(* IEC 61131-3 sources: plc-st-coding-agent/progress/evidence/v13_rescore_20261108/candidates/codex_minimax-m27, 19 files *)

(* ---- public-easy-01.st ---- *)
FUNCTION_BLOCK FB
VAR_INPUT
    bottleSensor           : BOOL;
    cleaningConfirmButton  : BOOL;
    fillingConfirmButton   : BOOL;
    cappingConfirmButton   : BOOL;
    packingConfirmButton   : BOOL;
    finishedButton         : BOOL;
END_VAR

VAR_OUTPUT
    Pump_Motor        : BOOL;
    Filling_Valve     : BOOL;
    Capping_Machine   : BOOL;
    Packing_Machine   : BOOL;
    Completion_Light  : BOOL;
END_VAR

VAR
    step                  : INT := 0;
    prevBottleSensor      : BOOL := FALSE;
    prevCleaningConfirm   : BOOL := FALSE;
    prevFillingConfirm    : BOOL := FALSE;
    prevCappingConfirm    : BOOL := FALSE;
    prevPackingConfirm    : BOOL := FALSE;
    prevFinishedButton    : BOOL := FALSE;
END_VAR

// Rising edge detection
VAR
    bottleRising         : BOOL;
    cleaningRising       : BOOL;
    fillingRising        : BOOL;
    cappingRising        : BOOL;
    packingRising        : BOOL;
    finishedRising       : BOOL;
END_VAR

bottleRising       := bottleSensor        AND NOT prevBottleSensor;
cleaningRising     := cleaningConfirmButton  AND NOT prevCleaningConfirm;
fillingRising      := fillingConfirmButton   AND NOT prevFillingConfirm;
cappingRising      := cappingConfirmButton   AND NOT prevCappingConfirm;
packingRising      := packingConfirmButton   AND NOT prevPackingConfirm;
finishedRising     := finishedButton      AND NOT prevFinishedButton;

// State machine transitions
IF step = 0 THEN
    IF bottleRising THEN
        step := 1;
    END_IF
ELSIF step = 1 THEN
    IF cleaningRising THEN
        step := 2;
    END_IF
ELSIF step = 2 THEN
    IF fillingRising THEN
        step := 3;
    END_IF
ELSIF step = 3 THEN
    IF cappingRising THEN
        step := 4;
    END_IF
ELSIF step = 4 THEN
    IF packingRising THEN
        step := 5;
    END_IF
END_IF

// Output logic based on step
Pump_Motor       := (step >= 1);
Filling_Valve    := (step >= 2);
Capping_Machine  := (step >= 3);
Packing_Machine  := (step >= 4);
Completion_Light := (step >= 5);

// Reset on finishedButton rising only when in COMPLETE state
IF finishedRising AND (step = 5) THEN
    step := 0;
END_IF

// Update previous states
prevBottleSensor    := bottleSensor;
prevCleaningConfirm := cleaningConfirmButton;
prevFillingConfirm  := fillingConfirmButton;
prevCappingConfirm  := cappingConfirmButton;
prevPackingConfirm  := packingConfirmButton;
prevFinishedButton  := finishedButton;
END_FUNCTION_BLOCK

(* ---- public-easy-02.st ---- *)
FUNCTION_BLOCK FB
VAR_INPUT
END_VAR
VAR_OUTPUT
    hasChanged      : BOOL;
    hasRisingEdges  : BOOL;
    risingBits      : DWORD;
    noOfRisingBits  : USINT;
    hasFallingEdges : BOOL;
    fallingBits     : DWORD;
    noOfFallingBits : USINT;
END_VAR
VAR
    prevValue : DWORD := 0;
    bitCheck  : DWORD;
    i         : USINT;
END_VAR

// Calculate rising edges: current=1 AND previous=0
risingBits := value AND NOT prevValue;

// Calculate falling edges: current=0 AND previous=1
fallingBits := NOT value AND prevValue;

// Detect if value has changed
hasChanged := (value <> prevValue);

// Set edge flags based on bit streams
hasRisingEdges := (risingBits <> 0);
hasFallingEdges := (fallingBits <> 0);

// Count rising bits
noOfRisingBits := 0;
bitCheck := risingBits;
FOR i := 0 TO 31 DO
    IF (bitCheck AND 1) = 1 THEN
        noOfRisingBits := noOfRisingBits + 1;
    END_IF;
    bitCheck := SHR(bitCheck, 1);
END_FOR;

// Count falling bits
noOfFallingBits := 0;
bitCheck := fallingBits;
FOR i := 0 TO 31 DO
    IF (bitCheck AND 1) = 1 THEN
        noOfFallingBits := noOfFallingBits + 1;
    END_IF;
    bitCheck := SHR(bitCheck, 1);
END_FOR;

// Update history for next cycle
prevValue := value;
END_FUNCTION_BLOCK

(* ---- public-easy-03.st ---- *)
FUNCTION_BLOCK FB
VAR_INPUT
    Value       : REAL;
    hiLevel     : REAL;
    loLevel     : REAL;
    hystWindow  : REAL;
END_VAR
VAR_OUTPUT
    hiAlarm     : BOOL;
    loAlarm     : BOOL;
    error       : BOOL;
    status      : WORD;
END_VAR

    // Parameter validation errors take priority
    IF loLevel >= hiLevel THEN
        error   := TRUE;
        status  := 16#8001;
        RETURN;
    END_IF

    IF hystWindow >= (hiLevel - loLevel) THEN
        error   := TRUE;
        status  := 16#8002;
        RETURN;
    END_IF

    // No error
    error  := FALSE;
    status := 16#0000;

    // High alarm with hysteresis
    // Trigger: Value > hiLevel
    // Reset:   Value < hiLevel - hystWindow
    IF Value > hiLevel THEN
        hiAlarm := TRUE;
    ELSIF Value < (hiLevel - hystWindow) THEN
        hiAlarm := FALSE;
    END_IF

    // Low alarm with hysteresis
    // Trigger: Value < loLevel
    // Reset:   Value > loLevel + hystWindow
    IF Value < loLevel THEN
        loAlarm := TRUE;
    ELSIF Value > (loLevel + hystWindow) THEN
        loAlarm := FALSE;
    END_IF

END_FUNCTION_BLOCK

(* ---- public-easy-04.st ---- *)
FUNCTION_BLOCK FB
VAR_INPUT
    VISCOSITY_OK     : BOOL;
    PASTE_E_STOP_NC  : BOOL;
    DebounceTime     : TIME;
    CycleTime        : TIME;
END_VAR
VAR_OUTPUT
    VFD_RUN          : BOOL;
    PUMP_MAINT_DUE   : BOOL;
    PUMP_RUNTIME_ACC : LINT;
END_VAR
VAR
    visc_debounce_acc : TIME := T#0s;
    visc_valid        : BOOL := FALSE;
END_VAR

// Debounce logic for viscosity condition
IF NOT VISCOSITY_OK THEN
    visc_debounce_acc := T#0s;
    visc_valid        := FALSE;
ELSIF visc_debounce_acc < DebounceTime THEN
    visc_debounce_acc := visc_debounce_acc + CycleTime;
    IF visc_debounce_acc >= DebounceTime THEN
        visc_debounce_acc := DebounceTime;
        visc_valid        := TRUE;
    END_IF
END_IF;

// VFD run permissive: E-STOP must be closed AND viscosity debounced valid
VFD_RUN := PASTE_E_STOP_NC AND visc_valid;

// Accumulate runtime (in hours) only while pump is running
IF VFD_RUN THEN
    PUMP_RUNTIME_ACC := PUMP_RUNTIME_ACC + TO_LINT(TIME_TO_INT(CycleTime) / 3600000);
END_IF;

// Maintenance due indication at 500 hours
PUMP_MAINT_DUE := (PUMP_RUNTIME_ACC >= 500);
END_FUNCTION_BLOCK

(* ---- public-easy-05.st ---- *)
FUNCTION_BLOCK FB
VAR_INPUT
    Gap_Exceeded : BOOL;
    Weld_E_Stop_NC : BOOL;
    DebounceTime : TIME;
END_VAR
VAR_OUTPUT
    Operator_Alert : BOOL;
    Weld_Soft_Start_Active : BOOL;
END_VAR
VAR
    init_cycle_count : INT := 5;
    gap_exceeded_prev : BOOL := FALSE;
    debounce_counter : INT := 0;
    debounce_required : INT := 50;
END_VAR

// Emergency stop priority - immediate reset regardless of state
IF NOT Weld_E_Stop_NC THEN
    Operator_Alert := FALSE;
    debounce_counter := 0;
    Weld_Soft_Start_Active := FALSE;
    gap_exceeded_prev := Gap_Exceeded;
    RETURN;
END_IF;

// Power-up initialization inhibition (5 scan cycles)
IF init_cycle_count > 0 THEN
    init_cycle_count := init_cycle_count - 1;
    Weld_Soft_Start_Active := TRUE;
    Operator_Alert := FALSE;
    debounce_counter := 0;
    gap_exceeded_prev := Gap_Exceeded;
    RETURN;
END_IF;

Weld_Soft_Start_Active := FALSE;
gap_exceeded_prev := Gap_Exceeded;

// Gap monitoring with debounce
IF Gap_Exceeded THEN
    debounce_counter := debounce_counter + 1;
    IF debounce_counter >= debounce_required THEN
        Operator_Alert := TRUE;
    ELSE
        Operator_Alert := FALSE;
    END_IF;
ELSE
    debounce_counter := 0;
    Operator_Alert := FALSE;
END_IF;
END_FUNCTION_BLOCK

(* ---- public-easy-06.st ---- *)
FUNCTION_BLOCK FB
VAR_INPUT
    DO_LOW : BOOL;
    AERATION_E_STOP_NC : BOOL;
END_VAR
VAR_OUTPUT
    BLOWER_RUN : BOOL;
    AERATION_BLOWER_CYCLE_COUNT : UINT;
END_VAR
VAR
    prev_blower_run : BOOL := FALSE;
    delay_counter : UINT := 0;
END_VAR

IF DO_LOW AND AERATION_E_STOP_NC THEN
    IF delay_counter < 5 THEN
        delay_counter := delay_counter + 1;
    END_IF
    IF delay_counter >= 5 THEN
        BLOWER_RUN := TRUE;
    ELSE
        BLOWER_RUN := FALSE;
    END_IF
ELSE
    BLOWER_RUN := FALSE;
    delay_counter := 0;
END_IF

IF BLOWER_RUN AND NOT prev_blower_run THEN
    AERATION_BLOWER_CYCLE_COUNT := AERATION_BLOWER_CYCLE_COUNT + 1;
END_IF

prev_blower_run := BLOWER_RUN;
END_FUNCTION_BLOCK

(* ---- public-hard-01.st ---- *)
FUNCTION_BLOCK FB
VAR_INPUT
    estop            : BOOL;
    opeMode          : BOOL;
    valveAStart      : BOOL;
    valveBStart      : BOOL;
    valveCStart      : BOOL;
    valveDStart      : BOOL;
    mixMotorStart    : BOOL;
    autoStart        : BOOL;
    processMode      : BOOL;
    levelSensor      : INT;
    mixMotorComplete : BOOL;
END_VAR
VAR_OUTPUT
    valveARun    : BOOL;
    valveBRun    : BOOL;
    valveCRun    : BOOL;
    valveDRun    : BOOL;
    mixMotorRun  : BOOL;
END_VAR
VAR
    // Auto mode state machine
    autoState : INT;
    // Rising edge detection history
    prevValveAStart    : BOOL;
    prevValveBStart    : BOOL;
    prevValveCStart    : BOOL;
    prevValveDStart    : BOOL;
    prevMixMotorStart  : BOOL;
    prevAutoStart      : BOOL;
    // Rising edge results
    valveAStartEdge    : BOOL;
    valveBStartEdge    : BOOL;
    valveCStartEdge    : BOOL;
    valveDStartEdge    : BOOL;
    mixMotorStartEdge  : BOOL;
    autoStartEdge      : BOOL;
END_VAR

    // Auto state constants
    // 0=IDLE, 1=VALVE_A, 2=VALVE_B, 3=VALVE_C, 4=MIXING, 5=DISCHARGE

    // Rising edge detection
    valveAStartEdge   := valveAStart AND NOT prevValveAStart;
    valveBStartEdge   := valveBStart AND NOT prevValveBStart;
    valveCStartEdge   := valveCStart AND NOT prevValveCStart;
    valveDStartEdge   := valveDStart AND NOT prevValveDStart;
    mixMotorStartEdge := mixMotorStart AND NOT prevMixMotorStart;
    autoStartEdge     := autoStart AND NOT prevAutoStart;

    // Update edge detection history
    prevValveAStart   := valveAStart;
    prevValveBStart   := valveBStart;
    prevValveCStart   := valveCStart;
    prevValveDStart   := valveDStart;
    prevMixMotorStart := mixMotorStart;
    prevAutoStart     := autoStart;

    // Default outputs off (safety)
    valveARun   := FALSE;
    valveBRun   := FALSE;
    valveCRun   := FALSE;
    valveDRun   := FALSE;
    mixMotorRun := FALSE;

    // Emergency stop - all equipment stops immediately
    IF NOT estop THEN
        autoState := 0;
        RETURN;
    END_IF

    // Manual mode
    IF NOT opeMode THEN
        // Rising edge toggles for each device
        IF valveAStartEdge THEN
            valveARun := NOT valveARun;
        END_IF
        IF valveBStartEdge THEN
            valveBRun := NOT valveBRun;
        END_IF
        IF valveCStartEdge THEN
            valveCRun := NOT valveCRun;
        END_IF
        IF valveDStartEdge THEN
            valveDRun := NOT valveDRun;
        END_IF
        IF mixMotorStartEdge THEN
            mixMotorRun := NOT mixMotorRun;
        END_IF
    // Automatic mode
    ELSIF opeMode THEN
        CASE autoState OF
            0: // IDLE
                IF autoStartEdge THEN
                    autoState := 1;
                END_IF

            1: // Open Valve A
                valveARun := TRUE;
                IF levelSensor >= 50 THEN
                    valveARun := FALSE;
                    autoState := 2;
                END_IF

            2: // Open Valve B
                valveBRun := TRUE;
                IF levelSensor >= 80 THEN
                    valveBRun := FALSE;
                    IF processMode THEN
                        autoState := 3;
                    ELSE
                        autoState := 4;
                    END_IF;
                END_IF

            3: // Open Valve C (processMode=true)
                valveCRun := TRUE;
                IF levelSensor >= 100 THEN
                    valveCRun := FALSE;
                    autoState := 4;
                END_IF

            4: // Mixing
                mixMotorRun := TRUE;
                IF mixMotorComplete THEN
                    mixMotorRun := FALSE;
                    autoState := 5;
                END_IF

            5: // Discharge through Valve D
                valveDRun := TRUE;
                IF levelSensor <= 0 THEN
                    valveDRun := FALSE;
                    autoState := 0;
                END_IF
        END_CASE
    END_IF

END_FUNCTION_BLOCK

(* ---- public-hard-02.st ---- *)
FUNCTION_BLOCK FB
VAR_INPUT
    processLength : USINT;
    sensor1 : BOOL;
    sensor2 : BOOL;
    sensor3 : BOOL;
    sensor4 : BOOL;
    sensor5 : BOOL;
    station1Start : BOOL;
    station2Complete : BOOL;
    station3Complete : BOOL;
    station4Complete : BOOL;
    processSequence : ARRAY[1..8] OF USINT;
END_VAR

VAR_OUTPUT
    conveyorLeft : BOOL;
    conveyorRight : BOOL;
END_VAR

VAR
    phase : USINT := 0;
    curStation : USINT := 0;
    dstStation : USINT := 0;
    idx : USINT := 1;
    prevStart : BOOL := FALSE;
    prevComp2 : BOOL := FALSE;
    prevComp3 : BOOL := FALSE;
    prevComp4 : BOOL := FALSE;
END_VAR

VAR
    startEdge : BOOL;
    compEdge : BOOL;
END_VAR

startEdge := station1Start AND NOT prevStart;
compEdge := (station2Complete AND NOT prevComp2) OR
            (station3Complete AND NOT prevComp3) OR
            (station4Complete AND NOT prevComp4);

prevStart := station1Start;
prevComp2 := station2Complete;
prevComp3 := station3Complete;
prevComp4 := station4Complete;

IF sensor1 AND startEdge THEN
    phase := 0;
    idx := 1;
    curStation := 1;
END_IF

CASE phase OF
    0:
        conveyorLeft := FALSE;
        conveyorRight := FALSE;
        IF sensor1 AND startEdge THEN
            curStation := 1;
            idx := 1;
            dstStation := processSequence[idx];
            phase := 1;
        END_IF

    1:
        IF dstStation > curStation THEN
            conveyorRight := TRUE;
            conveyorLeft := FALSE;
        ELSIF dstStation < curStation THEN
            conveyorLeft := TRUE;
            conveyorRight := FALSE;
        END_IF

        IF (dstStation = 2 AND sensor2) OR
           (dstStation = 3 AND sensor3) OR
           (dstStation = 4 AND sensor4) OR
           (dstStation = 5 AND sensor5) THEN
            curStation := dstStation;
            conveyorLeft := FALSE;
            conveyorRight := FALSE;
            phase := 2;
        END_IF

    2:
        conveyorLeft := FALSE;
        conveyorRight := FALSE;

        IF compEdge THEN
            IF curStation = 2 THEN
                idx := idx + 1;
                IF idx <= processLength THEN
                    dstStation := processSequence[idx];
                    phase := 1;
                END_IF
            ELSIF curStation = 3 THEN
                idx := idx + 1;
                IF idx <= processLength THEN
                    dstStation := processSequence[idx];
                    phase := 1;
                END_IF
            ELSIF curStation = 4 THEN
                idx := idx + 1;
                IF idx <= processLength THEN
                    dstStation := processSequence[idx];
                    phase := 1;
                END_IF
            END_IF
        END_IF

        IF curStation = 5 THEN
            phase := 0;
        END_IF
END_CASE
END_FUNCTION_BLOCK

(* ---- public-hard-03.st ---- *)
TYPE ST_Recipe :
STRUCT
    recipeID : INT;
    ingredientType : INT;
    ingredientRatio : REAL;
    productionTemperature : REAL;
END_STRUCT
END_TYPE

FUNCTION_BLOCK FB
VAR_INPUT
    addRecipe : BOOL;
    deleteRecipe : BOOL;
    modifyRecipe : BOOL;
    queryRecipe : BOOL;
    recipeIn : ST_Recipe;
END_VAR

VAR_OUTPUT
    recipeAdded : BOOL := FALSE;
    recipeDeleted : BOOL := FALSE;
    recipeModified : BOOL := FALSE;
    recipeQueryResult : ST_Recipe;
    error : BOOL := FALSE;
    status : WORD := 16#0000;
END_VAR

VAR_IN_OUT
    recipe : ARRAY[1..10] OF ST_Recipe;
END_VAR

VAR
    addRecipePrev : BOOL := FALSE;
    deleteRecipePrev : BOOL := FALSE;
    modifyRecipePrev : BOOL := FALSE;
    queryRecipePrev : BOOL := FALSE;
    foundIndex : INT;
    i : INT;
    isDuplicate : BOOL;
    isFound : BOOL;
END_VAR

    error := FALSE;
    status := 16#0000;
    recipeAdded := FALSE;
    recipeDeleted := FALSE;
    recipeModified := FALSE;

    IF addRecipe AND NOT addRecipePrev THEN
        isDuplicate := FALSE;
        isFound := FALSE;
        foundIndex := 0;

        FOR i := 1 TO 10 DO
            IF recipe[i].recipeID = recipeIn.recipeID AND recipeIn.recipeID <> 0 THEN
                isDuplicate := TRUE;
                EXIT;
            END_IF
        END_FOR

        IF isDuplicate THEN
            error := TRUE;
            status := 16#8002;
        ELSE
            foundIndex := 0;
            FOR i := 1 TO 10 DO
                IF recipe[i].recipeID = 0 THEN
                    foundIndex := i;
                    EXIT;
                END_IF
            END_FOR

            IF foundIndex = 0 THEN
                error := TRUE;
                status := 16#8003;
            ELSE
                recipe[foundIndex] := recipeIn;
                recipeAdded := TRUE;
            END_IF
        END_IF
    END_IF

    IF deleteRecipe AND NOT deleteRecipePrev THEN
        isFound := FALSE;
        foundIndex := 0;

        FOR i := 1 TO 10 DO
            IF recipe[i].recipeID = recipeIn.recipeID AND recipeIn.recipeID <> 0 THEN
                isFound := TRUE;
                foundIndex := i;
                EXIT;
            END_IF
        END_FOR

        IF NOT isFound THEN
            error := TRUE;
            status := 16#8004;
        ELSE
            recipe[foundIndex].recipeID := 0;
            recipeDeleted := TRUE;
        END_IF
    END_IF

    IF modifyRecipe AND NOT modifyRecipePrev THEN
        isFound := FALSE;
        foundIndex := 0;

        FOR i := 1 TO 10 DO
            IF recipe[i].recipeID = recipeIn.recipeID AND recipeIn.recipeID <> 0 THEN
                isFound := TRUE;
                foundIndex := i;
                EXIT;
            END_IF
        END_FOR

        IF NOT isFound THEN
            error := TRUE;
            status := 16#8005;
        ELSE
            recipe[foundIndex] := recipeIn;
            recipeModified := TRUE;
        END_IF
    END_IF

    IF queryRecipe AND NOT queryRecipePrev THEN
        isFound := FALSE;
        foundIndex := 0;

        FOR i := 1 TO 10 DO
            IF recipe[i].recipeID = recipeIn.recipeID AND recipeIn.recipeID <> 0 THEN
                isFound := TRUE;
                foundIndex := i;
                EXIT;
            END_IF
        END_FOR

        IF NOT isFound THEN
            error := TRUE;
            status := 16#8001;
        ELSE
            recipeQueryResult := recipe[foundIndex];
        END_IF
    END_IF

    addRecipePrev := addRecipe;
    deleteRecipePrev := deleteRecipe;
    modifyRecipePrev := modifyRecipe;
    queryRecipePrev := queryRecipe;

END_FUNCTION_BLOCK

(* ---- public-hard-04.st ---- *)
FUNCTION_BLOCK FB
VAR_INPUT
    enqueue  : BOOL;
    dequeue  : BOOL;
    reset    : BOOL;
    capacity : DINT;
END_VAR
VAR_OUTPUT
    elementCount : DINT := 0;
    status       : WORD := 16#0000;
END_VAR
VAR_IN_OUT
    item   : DINT;
    buffer : ARRAY[1..4] OF DINT;
END_VAR
VAR
    head        : DINT := 1;
    tail        : DINT := 1;
    lastEnqueue : BOOL := FALSE;
    lastDequeue : BOOL := FALSE;
    lastReset   : BOOL := FALSE;
END_VAR

status := 16#0000;

IF reset THEN
    elementCount := 0;
    head := 1;
    tail := 1;
ELSIF NOT lastReset THEN
    IF enqueue AND NOT lastEnqueue THEN
        IF elementCount < capacity THEN
            buffer[tail] := item;
            elementCount := elementCount + 1;
            tail := (tail MOD capacity) + 1;
        ELSE
            status := 16#8002;
        END_IF
    ELSIF dequeue AND NOT lastDequeue THEN
        IF elementCount > 0 THEN
            item := buffer[head];
            elementCount := elementCount - 1;
            head := (head MOD capacity) + 1;
        ELSE
            status := 16#8001;
        END_IF
    END_IF
END_IF

lastEnqueue := enqueue;
lastDequeue := dequeue;
lastReset   := reset;
END_FUNCTION_BLOCK

(* ---- public-hard-05.st ---- *)
FUNCTION_BLOCK FB
VAR_INPUT
    ManualMode : BOOL;
    SingleStepMode : BOOL;
    SingleCycleMode : BOOL;
    ContinuousMode : BOOL;
    EmergencyStop : BOOL;
    Start : BOOL;
    DownButton : BOOL;
    UpButton : BOOL;
    LeftButton : BOOL;
    RightButton : BOOL;
    GripButton : BOOL;
    ReleaseButton : BOOL;
    DownLimitSwitch : BOOL;
    UpLimitSwitch : BOOL;
    LeftLimitSwitch : BOOL;
    RightLimitSwitch : BOOL;
    GripLimitSwitch : BOOL;
    ReleaseLimitSwitch : BOOL;
END_VAR

VAR_OUTPUT
    MoveDown : BOOL := FALSE;
    MoveUp : BOOL := FALSE;
    MoveLeft : BOOL := FALSE;
    MoveRight : BOOL := FALSE;
    ActivateGrip : BOOL := FALSE;
    ActivateRelease : BOOL := FALSE;
END_VAR

VAR
    Step : INT := 1;
    StartPrev : BOOL := FALSE;
    IsRunning : BOOL := FALSE;
END_VAR

    // Edge detection for Start button
    VAR
        StartRisingEdge : BOOL;
    END_VAR
    StartRisingEdge := Start AND NOT StartPrev;
    StartPrev := Start;

    // Emergency stop - highest priority
    IF NOT EmergencyStop THEN
        MoveDown := FALSE;
        MoveUp := FALSE;
        MoveLeft := FALSE;
        MoveRight := FALSE;
        ActivateGrip := FALSE;
        ActivateRelease := FALSE;
        RETURN;
    END_IF

    // Mode initialization
    IF SingleStepMode THEN
        IF NOT IsRunning THEN
            IF StartRisingEdge THEN
                Step := 1;
                IsRunning := TRUE;
            END_IF;
        END_IF;
    ELSIF SingleCycleMode THEN
        IF NOT IsRunning THEN
            IF StartRisingEdge THEN
                Step := 1;
                IsRunning := TRUE;
            END_IF;
        END_IF;
    ELSIF ContinuousMode THEN
        IF NOT IsRunning THEN
            IF StartRisingEdge THEN
                Step := 1;
                IsRunning := TRUE;
            END_IF;
        END_IF;
    ELSE
        IsRunning := FALSE;
    END_IF;

    // Execute current step in automatic modes
    IF IsRunning THEN
        CASE Step OF
            1: // MoveDown
                MoveDown := TRUE;
                IF DownLimitSwitch THEN
                    MoveDown := FALSE;
                    IF Step < 8 THEN
                        Step := Step + 1;
                    ELSE
                        Step := 1;
                    END_IF;
                    IF SingleStepMode THEN
                        IsRunning := FALSE;
                    END_IF;
                END_IF;

            2: // ActivateGrip
                ActivateGrip := TRUE;
                IF GripLimitSwitch THEN
                    ActivateGrip := FALSE;
                    IF Step < 8 THEN
                        Step := Step + 1;
                    ELSE
                        Step := 1;
                    END_IF;
                    IF SingleStepMode THEN
                        IsRunning := FALSE;
                    END_IF;
                END_IF;

            3: // MoveUp
                MoveUp := TRUE;
                IF UpLimitSwitch THEN
                    MoveUp := FALSE;
                    IF Step < 8 THEN
                        Step := Step + 1;
                    ELSE
                        Step := 1;
                    END_IF;
                    IF SingleStepMode THEN
                        IsRunning := FALSE;
                    END_IF;
                END_IF;

            4: // MoveRight
                MoveRight := TRUE;
                IF RightLimitSwitch THEN
                    MoveRight := FALSE;
                    IF Step < 8 THEN
                        Step := Step + 1;
                    ELSE
                        Step := 1;
                    END_IF;
                    IF SingleStepMode THEN
                        IsRunning := FALSE;
                    END_IF;
                END_IF;

            5: // MoveDown
                MoveDown := TRUE;
                IF DownLimitSwitch THEN
                    MoveDown := FALSE;
                    IF Step < 8 THEN
                        Step := Step + 1;
                    ELSE
                        Step := 1;
                    END_IF;
                    IF SingleStepMode THEN
                        IsRunning := FALSE;
                    END_IF;
                END_IF;

            6: // ActivateRelease
                ActivateRelease := TRUE;
                IF ReleaseLimitSwitch THEN
                    ActivateRelease := FALSE;
                    IF Step < 8 THEN
                        Step := Step + 1;
                    ELSE
                        Step := 1;
                    END_IF;
                    IF SingleStepMode THEN
                        IsRunning := FALSE;
                    END_IF;
                END_IF;

            7: // MoveUp
                MoveUp := TRUE;
                IF UpLimitSwitch THEN
                    MoveUp := FALSE;
                    IF Step < 8 THEN
                        Step := Step + 1;
                    ELSE
                        Step := 1;
                    END_IF;
                    IF SingleStepMode THEN
                        IsRunning := FALSE;
                    END_IF;
                END_IF;

            8: // MoveLeft
                MoveLeft := TRUE;
                IF LeftLimitSwitch THEN
                    MoveLeft := FALSE;
                    Step := 1;
                    IF SingleStepMode THEN
                        IsRunning := FALSE;
                    END_IF;
                END_IF;
        END_CASE;

    // Manual mode
    ELSIF ManualMode THEN
        // Down
        MoveDown := DownButton AND NOT DownLimitSwitch;
        // Up
        MoveUp := UpButton AND NOT UpLimitSwitch;
        // Left
        MoveLeft := LeftButton AND NOT LeftLimitSwitch;
        // Right
        MoveRight := RightButton AND NOT RightLimitSwitch;
        // Grip
        ActivateGrip := GripButton AND NOT GripLimitSwitch;
        // Release
        ActivateRelease := ReleaseButton AND NOT ReleaseLimitSwitch;
    END_IF;

END_FUNCTION_BLOCK

(* ---- public-hard-06.st ---- *)
FUNCTION_BLOCK FB
VAR_INPUT
    Mode            : BOOL;
    ForwardButton   : BOOL;
    ReverseButton   : BOOL;
    SensorFeed      : BOOL;
    SensorWash      : BOOL;
    SensorWeight    : BOOL;
    SensorFiring    : BOOL;
    SensorOutput    : BOOL;
    washComplete    : BOOL;
    weightComplete  : BOOL;
    weight          : REAL;
    firingComplete  : BOOL;
END_VAR
VAR_OUTPUT
    MotorForward    : BOOL;
    MotorReverse    : BOOL;
    kick            : BOOL;
    CompletionLight : BOOL;
    firingTemp      : REAL;
END_VAR
VAR
    eState              : INT;
    prevForwardButton   : BOOL;
    prevReverseButton   : BOOL;
    prevwashComplete    : BOOL;
    prevweightComplete  : BOOL;
    prevfiringComplete  : BOOL;
    bKickDone           : BOOL;
END_VAR

    // Edge detection: rising edge flags
    VAR
        bFwdRising   : BOOL;
        bRevRising   : BOOL;
        bWashRising  : BOOL;
        bWeightRising: BOOL;
        bFiringRising: BOOL;
    END_VAR

    bFwdRising   := (NOT prevForwardButton)  AND ForwardButton;
    bRevRising   := (NOT prevReverseButton)  AND ReverseButton;
    bWashRising  := (NOT prevwashComplete)   AND washComplete;
    bWeightRising:= (NOT prevweightComplete) AND weightComplete;
    bFiringRising:= (NOT prevfiringComplete) AND firingComplete;

    // Reset kick flag on new cycle start (ForwardButton rising edge in any mode)
    IF bFwdRising THEN
        bKickDone := FALSE;
    END_IF

    IF Mode = FALSE THEN
        // Manual mode
        eState := 0;
        MotorForward := ForwardButton;
        MotorReverse := ReverseButton;
        kick := FALSE;
        CompletionLight := FALSE;
        firingTemp := 0.0;
    ELSE
        // Automatic mode
        CASE eState OF
            0:  // IDLE
                MotorForward := FALSE;
                MotorReverse := FALSE;
                kick := FALSE;
                CompletionLight := FALSE;
                firingTemp := 0.0;
                bKickDone := FALSE;
                IF SensorFeed THEN
                    eState := 1;
                END_IF

            1:  // MOVING_TO_WASH
                MotorForward := TRUE;
                MotorReverse := FALSE;
                kick := FALSE;
                IF SensorWash THEN
                    eState := 2;
                END_IF

            2:  // AT_WASH
                MotorForward := FALSE;
                MotorReverse := FALSE;
                kick := FALSE;
                IF bWashRising THEN
                    eState := 3;
                END_IF

            3:  // MOVING_TO_WEIGH
                MotorForward := TRUE;
                MotorReverse := FALSE;
                kick := FALSE;
                IF SensorWeight THEN
                    eState := 4;
                END_IF

            4:  // AT_WEIGH
                MotorForward := FALSE;
                MotorReverse := FALSE;
                kick := FALSE;
                IF bWeightRising THEN
                    IF weight >= 100.0 AND weight <= 200.0 THEN
                        firingTemp := 500.0 + (weight - 100.0) * 0.5;
                        eState := 6;
                    ELSE
                        eState := 5;
                    END_IF;
                END_IF

            5:  // KICKING
                MotorForward := FALSE;
                MotorReverse := FALSE;
                kick := TRUE;
                IF NOT bKickDone THEN
                    bKickDone := TRUE;
                    eState := 0;
                END_IF

            6:  // MOVING_TO_FIRING
                MotorForward := TRUE;
                MotorReverse := FALSE;
                kick := FALSE;
                IF SensorFiring THEN
                    eState := 7;
                END_IF

            7:  // AT_FIRING
                MotorForward := FALSE;
                MotorReverse := FALSE;
                kick := FALSE;
                IF bFiringRising THEN
                    eState := 8;
                END_IF

            8:  // MOVING_TO_OUTPUT
                MotorForward := TRUE;
                MotorReverse := FALSE;
                kick := FALSE;
                IF SensorOutput THEN
                    eState := 9;
                END_IF

            9:  // AT_OUTPUT
                MotorForward := FALSE;
                MotorReverse := FALSE;
                kick := FALSE;
                CompletionLight := SensorOutput;
                IF NOT SensorOutput THEN
                    eState := 0;
                END_IF

        END_CASE
    END_IF

    prevForwardButton  := ForwardButton;
    prevReverseButton  := ReverseButton;
    prevwashComplete   := washComplete;
    prevweightComplete := weightComplete;
    prevfiringComplete := firingComplete;

END_FUNCTION_BLOCK

(* ---- public-medium-01.st ---- *)
TYPE ST_Pump
    STRUCT
        priority   : INT;
        selection  : BOOL;
        RunComd    : BOOL;
    END_STRUCT
END_TYPE

FUNCTION_BLOCK FB
VAR_INPUT
    mode  : BOOL;
    start : BOOL;
    stop  : BOOL;
END_VAR
VAR_IN_OUT
    pumpGroup : ARRAY[1..5] OF ST_Pump;
END_VAR
VAR
    prevStart     : BOOL := FALSE;
    prevStop      : BOOL := FALSE;
    i             : INT;
    j             : INT;
    k             : INT;
    tmp           : INT;
    tmpIdx        : INT;
    tempPriority  : ARRAY[1..5] OF INT;
    sortedIdx     : ARRAY[1..5] OF INT;
END_VAR

IF stop THEN
    FOR i := 1 TO 5 DO
        pumpGroup[i].RunComd := FALSE;
    END_FOR;
ELSE
    IF start AND NOT prevStart THEN
        IF NOT mode THEN
            FOR i := 1 TO 5 DO
                IF pumpGroup[i].selection THEN
                    pumpGroup[i].RunComd := TRUE;
                ELSE
                    pumpGroup[i].RunComd := FALSE;
                END_IF;
            END_FOR;
        ELSE
            FOR i := 1 TO 5 DO
                tempPriority[i] := pumpGroup[i].priority;
                sortedIdx[i] := i;
            END_FOR;
            FOR j := 1 TO 4 DO
                FOR k := j + 1 TO 5 DO
                    IF tempPriority[k] > tempPriority[j] OR
                       (tempPriority[k] = tempPriority[j] AND sortedIdx[k] < sortedIdx[j]) THEN
                        tmp := tempPriority[j];
                        tempPriority[j] := tempPriority[k];
                        tempPriority[k] := tmp;
                        tmpIdx := sortedIdx[j];
                        sortedIdx[j] := sortedIdx[k];
                        sortedIdx[k] := tmpIdx;
                    END_IF;
                END_FOR;
            END_FOR;
            FOR i := 1 TO 5 DO
                IF i <= 3 THEN
                    pumpGroup[sortedIdx[i]].RunComd := TRUE;
                ELSE
                    pumpGroup[sortedIdx[i]].RunComd := FALSE;
                END_IF;
            END_FOR;
        END_IF;
    ELSE
        FOR i := 1 TO 5 DO
            pumpGroup[i].RunComd := FALSE;
        END_FOR;
    END_IF;
END_IF;

prevStart := start;
prevStop := stop;

END_FUNCTION_BLOCK

(* ---- public-medium-02.st ---- *)
TYPE ST_AnalogChannel :
STRUCT
    enable       : BOOL;
    hiLIM        : REAL;
    loLIM        : REAL;
    bipolar      : BOOL;
    measuringMode: INT;
    retVal       : WORD;
    outputValue  : REAL;
END_STRUCT
END_TYPE

FUNCTION_BLOCK FB
VAR_INPUT
    count : DINT;
END_VAR
VAR_IN_OUT
    analogValues : ARRAY[1..8] OF INT;
    channels     : ARRAY[1..8] OF ST_AnalogChannel;
END_VAR
VAR
    i   : DINT;
    raw : INT;
END_VAR

IF count < 1 THEN
    RETURN;
END_IF;

FOR i := 1 TO count DO
    IF channels[i].enable THEN
        raw := analogValues[i];

        IF channels[i].measuringMode < 0 OR channels[i].measuringMode > 2 THEN
            channels[i].retVal := 16#8001;
        ELSIF channels[i].hiLIM <= channels[i].loLIM THEN
            channels[i].retVal := 16#8002;
        ELSIF channels[i].measuringMode = 0 THEN
            IF NOT channels[i].bipolar THEN
                channels[i].outputValue := channels[i].loLIM
                    + (INT_TO_REAL(raw) / 27648.0)
                    * (channels[i].hiLIM - channels[i].loLIM);
            ELSE
                channels[i].outputValue := channels[i].loLIM
                    + ((INT_TO_REAL(raw) + 27648.0) / (2.0 * 27648.0))
                    * (channels[i].hiLIM - channels[i].loLIM);
            END_IF;
            channels[i].retVal := 16#0000;
        ELSIF channels[i].measuringMode = 1 THEN
            channels[i].outputValue := INT_TO_REAL(raw) / 10.0;
            channels[i].retVal      := 16#0000;
        ELSIF channels[i].measuringMode = 2 THEN
            channels[i].outputValue := INT_TO_REAL(raw) / 100.0;
            channels[i].retVal      := 16#0000;
        END_IF;
    END_IF;
END_FOR
END_FUNCTION_BLOCK

(* ---- public-medium-03.st ---- *)
FUNCTION_BLOCK FB
VAR_INPUT
    cyclicExecution : BOOL;
    trigger : BOOL;
    value : LREAL;
    windowSize : INT;
    reset : BOOL;
END_VAR

VAR_OUTPUT
    average : LREAL := 0.0;
    windowSizeReached : BOOL := FALSE;
    error : BOOL := FALSE;
    status : WORD := 16#0000;
END_VAR

VAR
    dataBuffer : ARRAY[1..100] OF LREAL;
    sampleCount : INT := 0;
    nextIndex : INT := 1;
    lastTrigger : BOOL := FALSE;
    sum : LREAL;
    i : INT;
END_VAR

// Reset on rising edge when no error
IF reset AND NOT error THEN
    sampleCount := 0;
    nextIndex := 1;
    average := 0.0;
    windowSizeReached := FALSE;
END_IF

// Window size validation
IF (windowSize < 1) OR (windowSize > 100) THEN
    error := TRUE;
    status := 16#8200;
    IF error THEN
        RETURN;
    END_IF
END_IF

// Clear error when window size becomes valid
IF NOT error THEN
    error := FALSE;
    status := 16#0000;
END_IF

// Handle cyclic or trigger-based updates
IF cyclicExecution OR (trigger AND NOT lastTrigger) THEN
    IF sampleCount < windowSize THEN
        sampleCount := sampleCount + 1;
        dataBuffer[sampleCount] := value;
    ELSE
        dataBuffer[nextIndex] := value;
        nextIndex := (nextIndex MOD windowSize) + 1;
    END_IF

    // Recalculate average
    sum := 0.0;
    FOR i := 1 TO sampleCount DO
        sum := sum + dataBuffer[i];
    END_FOR
    average := sum / INT_TO_LREAL(sampleCount);
END_IF

// Update window size reached flag
windowSizeReached := (sampleCount >= windowSize);

// Update lastTrigger
lastTrigger := trigger;

END_FUNCTION_BLOCK

(* ---- public-medium-04.st ---- *)
FUNCTION_BLOCK FB
VAR_INPUT
    TemperatureSensorInput : REAL;
    SetTemperature : REAL;
END_VAR
VAR_OUTPUT
    CurrentTemperature : REAL;
    SetTempDisplay : REAL;
    HeaterStatus : BOOL;
    OverheatProtection : BOOL;
    HeaterOutput : BOOL;
END_VAR
VAR
    ContinuousHeatingCount : INT := 0;
    OverheatProtectionCount : INT := 0;
    PrevHeaterOutput : BOOL := FALSE;
END_VAR

// Determine if sensor has a fault
IF TemperatureSensorInput < 0.0 OR TemperatureSensorInput > 100.0 THEN
    // Sensor fault - turn off heater
    HeaterOutput := FALSE;
    ContinuousHeatingCount := 0;
ELSE
    // No sensor fault - check overheat protection status
    IF OverheatProtection THEN
        // Overheat protection is active
        HeaterOutput := FALSE;
        ContinuousHeatingCount := 0;

        // Overheat protection can only be cleared after 3 cycles
        IF PrevHeaterOutput = FALSE THEN
            OverheatProtectionCount := OverheatProtectionCount + 1;
            IF OverheatProtectionCount >= 3 THEN
                OverheatProtection := FALSE;
                OverheatProtectionCount := 0;
            END_IF
        END_IF
    ELSE
        // No overheat protection - normal temperature control
        IF TemperatureSensorInput < SetTemperature THEN
            // Temperature below set value - start heater
            HeaterOutput := TRUE;
        ELSE
            // Temperature at or above set value - stop heater
            HeaterOutput := FALSE;
        END_IF

        OverheatProtectionCount := 0;

        // Track continuous heating time (1 cycle = 1 second)
        IF HeaterOutput THEN
            ContinuousHeatingCount := ContinuousHeatingCount + 1;
            // Trigger overheat protection after 5 seconds continuous heating
            IF ContinuousHeatingCount >= 5 THEN
                OverheatProtection := TRUE;
                HeaterOutput := FALSE;
                ContinuousHeatingCount := 0;
            END_IF
        ELSE
            ContinuousHeatingCount := 0;
        END_IF
    END_IF
END_IF

// Update status outputs
CurrentTemperature := TemperatureSensorInput;
SetTempDisplay := SetTemperature;
HeaterStatus := HeaterOutput;

// Update previous heater output for edge detection
PrevHeaterOutput := HeaterOutput;
END_FUNCTION_BLOCK

(* ---- public-medium-05.st ---- *)
FUNCTION_BLOCK FB
VAR_INPUT
    Mode            : BOOL;
    ForwardButton   : BOOL;
    ReverseButton   : BOOL;
    SensorA         : BOOL;
    SensorB         : BOOL;
    SensorC         : BOOL;
    ButtonA         : BOOL;
    ButtonB         : BOOL;
    ButtonC         : BOOL;
END_VAR
VAR_OUTPUT
    MotorForward    : BOOL;
    MotorReverse    : BOOL;
    CompletionLight : BOOL;
END_VAR
VAR
    State           : INT := 0;
    prevSensorA     : BOOL := FALSE;
    prevSensorB     : BOOL := FALSE;
    prevSensorC     : BOOL := FALSE;
    prevButtonA     : BOOL := FALSE;
    prevButtonB     : BOOL := FALSE;
    prevButtonC     : BOOL := FALSE;
    SensorARising   : BOOL;
    SensorBRising   : BOOL;
    SensorCRising   : BOOL;
    ButtonARising   : BOOL;
    ButtonBRising   : BOOL;
    ButtonCRising   : BOOL;
END_VAR

// Edge detection
ButtonARising := ButtonA AND NOT prevButtonA;
ButtonBRising := ButtonB AND NOT prevButtonB;
ButtonCRising := ButtonC AND NOT prevButtonC;
SensorARising := SensorA AND NOT prevSensorA;
SensorBRising := SensorB AND NOT prevSensorB;
SensorCRising := SensorC AND NOT prevSensorC;

// Update history
prevButtonA := ButtonA;
prevButtonB := ButtonB;
prevButtonC := ButtonC;
prevSensorA := SensorA;
prevSensorB := SensorB;
prevSensorC := SensorC;

// Initialize outputs
MotorForward    := FALSE;
MotorReverse    := FALSE;
CompletionLight := FALSE;

// Automatic mode state machine
IF Mode THEN
    CASE State OF
        0: // IDLE
            IF SensorARising THEN
                State := 1;
            END_IF

        1: // WAIT_A
            MotorForward := FALSE;
            IF ButtonARising THEN
                State := 2;
            END_IF

        2: // Moving A->B
            MotorForward := TRUE;
            IF SensorBRising THEN
                State := 3;
            END_IF

        3: // WAIT_B
            MotorForward := FALSE;
            IF ButtonBRising THEN
                State := 4;
            END_IF

        4: // Moving B->C
            MotorForward := TRUE;
            IF SensorCRising THEN
                State := 5;
            END_IF

        5: // WAIT_C
            MotorForward := FALSE;
            CompletionLight := SensorC;
            IF NOT SensorC THEN
                State := 0;
            END_IF
    END_CASE
ELSE
    // Manual mode: reset state and handle interlocked control
    State := 0;

    IF ForwardButton AND NOT ReverseButton THEN
        MotorForward := TRUE;
    ELSIF ReverseButton AND NOT ForwardButton THEN
        MotorReverse := TRUE;
    END_IF
END_IF
END_FUNCTION_BLOCK

(* ---- public-medium-06.st ---- *)
FUNCTION_BLOCK FB
VAR_INPUT
    THICKNESS_FAULT        : BOOL;
    THICKNESS_SIGNAL_VALID : BOOL;
    CUTTING_RUN            : BOOL;
    FaultTimestamp         : DINT;
    CycleTime              : TIME;
END_VAR
VAR_OUTPUT
    THICKNESS_ALARM           : BOOL := FALSE;
    Slab_Fault_Counter        : UINT := 0;
    Slab_Runtime_Accumulator  : LINT := 0;
    Slab_Fault_History        : ARRAY[0..4] OF DINT;
END_VAR
VAR
    FaultPrev      : BOOL := FALSE;
    AlarmHoldTimer : TON;
    i              : INT;
END_VAR

    IF NOT THICKNESS_SIGNAL_VALID THEN
        THICKNESS_ALARM := FALSE;
        Slab_Fault_Counter := 0;
        Slab_Runtime_Accumulator := 0;
        Slab_Fault_History[0] := 0;
        Slab_Fault_History[1] := 0;
        Slab_Fault_History[2] := 0;
        Slab_Fault_History[3] := 0;
        Slab_Fault_History[4] := 0;
        AlarmHoldTimer(IN := FALSE);
        FaultPrev := FALSE;
    ELSE
        IF THICKNESS_FAULT THEN
            AlarmHoldTimer(IN := TRUE, PT := T#500ms);
            IF NOT FaultPrev THEN
                Slab_Fault_Counter := Slab_Fault_Counter + 1;
                FOR i := 4 TO 1 BY -1 DO
                    Slab_Fault_History[i] := Slab_Fault_History[i-1];
                END_FOR;
                Slab_Fault_History[0] := FaultTimestamp;
            END_IF;
        ELSE
            AlarmHoldTimer(IN := FALSE);
        END_IF;
        IF CUTTING_RUN THEN
            Slab_Runtime_Accumulator := Slab_Runtime_Accumulator + TIME_TO_LINT(CycleTime);
        END_IF;
        THICKNESS_ALARM := THICKNESS_FAULT OR AlarmHoldTimer.Q;
        FaultPrev := THICKNESS_FAULT;
    END_IF;

END_FUNCTION_BLOCK

(* ---- public-medium-07.st ---- *)
FUNCTION_BLOCK FB
VAR_INPUT
    OCCUPANCY_DETECTED    : BOOL;
    ENERGY_SAVING_MODE    : BOOL;
    HVAC_MODE_SELECTOR    : INT;
END_VAR

VAR_OUTPUT
    SUPPLY_FAN_RUN        : BOOL := FALSE;
    TEMP_SETPOINT_ADJUST  : INT  := 0;
END_VAR

VAR
    prev_start_condition  : BOOL := FALSE;
    delay_counter         : INT  := 0;
END_VAR

SUPPLY_FAN_RUN     := FALSE;
TEMP_SETPOINT_ADJUST := 0;

IF OCCUPANCY_DETECTED AND (HVAC_MODE_SELECTOR <> 3) THEN
    IF prev_start_condition THEN
        delay_counter := delay_counter + 1;
    ELSE
        delay_counter := 1;
    END_IF;
    IF delay_counter >= 30 THEN
        SUPPLY_FAN_RUN := TRUE;
    END_IF;
ELSE
    delay_counter := 0;
END_IF;
prev_start_condition := OCCUPANCY_DETECTED AND (HVAC_MODE_SELECTOR <> 3);

CASE HVAC_MODE_SELECTOR OF
    0:
        IF OCCUPANCY_DETECTED THEN
            TEMP_SETPOINT_ADJUST := 0;
        ELSIF ENERGY_SAVING_MODE THEN
            TEMP_SETPOINT_ADJUST := 3;
        ELSE
            TEMP_SETPOINT_ADJUST := 2;
        END_IF;
    1:
        IF OCCUPANCY_DETECTED THEN
            TEMP_SETPOINT_ADJUST := 0;
        ELSE
            TEMP_SETPOINT_ADJUST := 1;
        END_IF;
    2:
        IF OCCUPANCY_DETECTED THEN
            TEMP_SETPOINT_ADJUST := 0;
        ELSE
            TEMP_SETPOINT_ADJUST := 4;
        END_IF;
    3:
        TEMP_SETPOINT_ADJUST := 4;
ELSE
    TEMP_SETPOINT_ADJUST := 0;
END_CASE;

IF TEMP_SETPOINT_ADJUST < -4 THEN
    TEMP_SETPOINT_ADJUST := -4;
ELSIF TEMP_SETPOINT_ADJUST > 4 THEN
    TEMP_SETPOINT_ADJUST := 4;
END_IF;
END_FUNCTION_BLOCK
